Fanuc KAREL source: KA00100.KL

PROGRAM KA00100
%NOLOCKGROUP
VAR
  SRC: VECTOR
  DST: STRING[80]
BEGIN
  SRC.X = 1.0
  DST = SRC
END KA00100
